TEXTLIST TextList_Piston_Recipe_State_UpDown
  0 = ' '
  1 = 'Up'
  2 = 'Down'
   = ''
END_TEXTLIST

(* stored: Version 1.1.0.1, ProductVersion 3.1.4024.12
   TextList TextList_Piston_Recipe_State_UpDown: Id {ad52dd20-40d8-4d1b-8ecf-1cc30c39baf6} *)
